(*~
	<docu>
		<summary>
			Current test step (input 0Eh). None = FFFFh on the bus (no cycle running).
		</summary>
	</docu>
~*)
{attribute 'qualified_only'}
{attribute 'strict'}
TYPE eTcoAteqG6_Step_v_3_5_x :
(
	Unknown := -2,
	None := -1,
	PreFill := 0,
	Fill := 1,
	ZeroDiff := 2,
	Stabilization := 3,
	Test := 4,
	Dump := 5
) INT;
END_TYPE

(* stored: Version 1.1.0.1, ProductVersion 3.1.4024.12
   DUT eTcoAteqG6_Step_v_3_5_x: Id {620add64-f698-4724-9c8f-401a70abcc6d} *)
